TYPE "DT_PAR_PID_PELTON_NOZZLE_3"
VERSION : 0.1
   STRUCT
      INPUT_RAMP_MIN_VAL { S7_SetPoint := 'False'} : "DT_PARAM_SOLO" := (FALSE, 960, 0, 0.0, 0, T#0MS, 0.0, 0.0, '%');
      INPUT_RAMP_MAX_VAL { S7_SetPoint := 'False'} : "DT_PARAM_SOLO" := (FALSE, 961, 0, 100.0, 0, T#0MS, 0.0, 0.0, '%');
      INPUT_RAMP_FALLING_TIME { S7_SetPoint := 'False'} : "DT_PARAM_SOLO" := (FALSE, 962, 0, 0.0, 0, T#2M, 0.0, 0.0, 's');
      INPUT_RAMP_RISING_TIME { S7_SetPoint := 'False'} : "DT_PARAM_SOLO" := (FALSE, 963, 0, 0.0, 0, T#2M, 0.0, 0.0, 's');
      OUTPUT_RAMP_FALLING_TIME { S7_SetPoint := 'False'} : "DT_PARAM_SOLO" := (FALSE, 964, 0, 0.0, 0, T#0MS, 0.0, 0.0, 's');
      OUTPUT_RAMP_RISING_TIME { S7_SetPoint := 'False'} : "DT_PARAM_SOLO" := (FALSE, 965, 0, 0.0, 0, T#0MS, 0.0, 0.0, 's');
      MAN_ON { S7_SetPoint := 'False'} : "DT_PARAM_SOLO" := (FALSE, 966, 1, 0.0, 0, T#0MS, 0.0, 0.0, '-');
      P_SEL { S7_SetPoint := 'False'} : "DT_PARAM_SOLO" := (FALSE, 967, 1, 0.0, 1, T#0MS, 0.0, 0.0, '-');
      I_SEL { S7_SetPoint := 'False'} : "DT_PARAM_SOLO" := (FALSE, 968, 1, 0.0, 1, T#0MS, 0.0, 0.0, '-');
      INT_HOLD { S7_SetPoint := 'False'} : "DT_PARAM_SOLO" := (FALSE, 969, 1, 0.0, 0, T#0MS, 0.0, 0.0, '-');
      D_SEL { S7_SetPoint := 'False'} : "DT_PARAM_SOLO" := (FALSE, 970, 1, 0.0, 0, T#0MS, 0.0, 0.0, '-');
      NUM_OF_CYCLES { S7_SetPoint := 'False'} : "DT_PARAM_SOLO" := (FALSE, 971, 1, 0.0, 40, T#0MS, 0.0, 0.0, '-');
      GAIN { S7_SetPoint := 'False'} : "DT_PARAM_SOLO" := (FALSE, 972, 0, 13.0, 0, T#2M, 0.0, 0.0, '');
      TI { S7_SetPoint := 'False'} : "DT_PARAM_SOLO" := (FALSE, 973, 2, 0.0, 0, T#2M, 0.0, 0.0, '-');
      TD { S7_SetPoint := 'False'} : "DT_PARAM_SOLO" := (FALSE, 974, 2, 0.0, 0, T#0MS, 0.0, 0.0, '-');
      TM_LAG { S7_SetPoint := 'False'} : "DT_PARAM_SOLO" := (FALSE, 975, 2, 300.0, 0, T#0MS, 0.0, 0.0, '-');
      DEAD_W { S7_SetPoint := 'False'} : "DT_PARAM_SOLO" := (FALSE, 976, 0, 0.2, 0, T#2M, 0.0, 0.0, '%');
      LMN_HLM { S7_SetPoint := 'False'} : "DT_PARAM_SOLO" := (FALSE, 977, 0, 100.0, 0, T#0MS, 0.0, 0.0, '%');
      LMN_LLM { S7_SetPoint := 'False'} : "DT_PARAM_SOLO" := (FALSE, 978, 0, -100.0, 0, T#0MS, 0.0, 0.0, '%');
      REF_MIN_VAL { S7_SetPoint := 'False'} : "DT_PARAM_SOLO" := (FALSE, 979, 0, 0.0, 0, T#0MS, 0.0, 0.0, '%');
      REF_MAX_VAL { S7_SetPoint := 'False'} : "DT_PARAM_SOLO" := (FALSE, 980, 0, 100.0, 0, T#0MS, 0.0, 0.0, '%');
      LMN_FAC { S7_SetPoint := 'False'} : "DT_PARAM_SOLO" := (FALSE, 981, 0, 1.0, 0, T#0MS, 0.0, 0.0, '-');
      LMN_OFFSET { S7_SetPoint := 'False'} : "DT_PARAM_SOLO" := (FALSE, 982, 0, 0.0, 0, T#0MS, 0.0, 0.0, '%');
      DISV { S7_SetPoint := 'False'} : "DT_PARAM_SOLO" := (FALSE, 983, 0, 0.0, 0, T#0MS, 0.0, 0.0, '-');
      MAN { S7_SetPoint := 'False'} : "DT_PARAM_SOLO" := (FALSE, 984, 0, 0.0, 1, T#17S, 0.0, 0.0, '%');
      REFERENCE_CORRECTION { S7_SetPoint := 'False'} : "DT_PARAM_SOLO" := (FALSE, 985, 0, 0.0, 0, T#0MS, 0.0, 0.0, '-');
      OUT_CTRL_MODE { S7_SetPoint := 'False'} : "DT_PARAM_SOLO" := (FALSE, 986, 1, 0.0, 0, T#0MS, 0.0, 0.0, '-');
      SPARE_4 { S7_SetPoint := 'False'} : "DT_PARAM_SOLO" := (FALSE, 987, 0, 0.0, 0, T#0MS, 0.0, 0.0, '');
      SPARE_5 { S7_SetPoint := 'False'} : "DT_PARAM_SOLO" := (FALSE, 988, 0, 0.0, 0, T#0MS, 0.0, 0.0, '');
      SPARE_6 { S7_SetPoint := 'False'} : "DT_PARAM_SOLO" := (FALSE, 989, 0, 0.0, 0, T#0MS, 0.0, 0.0, '');
      SPARE_7 { S7_SetPoint := 'False'} : "DT_PARAM_SOLO" := (FALSE, 990, 0, 0.0, 0, T#0MS, 0.0, 0.0, '');
      SPARE_8 { S7_SetPoint := 'False'} : "DT_PARAM_SOLO" := (FALSE, 991, 0, 0.0, 0, T#0MS, 0.0, 0.0, '');
   END_STRUCT;

END_TYPE

